Fanuc KAREL source: kb00099.KL

-- PROVISIONAL review KL for V770-1; original PC SHA256 b27553b149da1b38c8a315ecbe82831e2fd5d384c5e63f24b1a36294e77b62be
-- Incomplete behavior may be omitted. Consult companion uncertainty JSON. Do not deploy.
PROGRAM KB00099
%NOLOCKGROUP
VAR
  P1 : STRING[80]
  P2 : STRING[80]
  RESULT : INTEGER
BEGIN
  -- UNRESOLVED_PC offsets 5-14; opcodes 3F,75
  -- UNRESOLVED_PC offsets 19-28; opcodes 3F,75
  -- UNRESOLVED_PC offsets 33-58; opcodes 27,22,2A,22,2A,76,23
  -- UNRESOLVED_PC offsets 63-67; opcodes 7F
END KB00099
